// TIA Portal V19 export
VAR_GLOBAL   // PLC tag table "Yaskawa_Inverter"
   INV_CMD AT %QW74 : Word;
   INV_CmdVelocity AT %QW76 : Word;
   INV_ETA AT %IW86 : Word;
   INV_ActRPM AT %IW88 : Word;
END_VAR
